Fanuc KAREL source: KT00708.KL

PROGRAM KT00708
%NOLOCKGROUP
VAR
  R1: REAL
  R2: REAL
  OUT: BOOLEAN
BEGIN
  R1 = 2.0
  R2 = 3.0
  R1 = 2.0
  R2 = 3.0
  OUT = UNINIT(R1)
END KT00708
